(* IEC 61131-3 sources: Lasal-MCP/examples/SampleSource/LASALScreenAdvancedSolution/LASALScreenAdvancedSolution/LASALScreenAdvacnedSolution/Stations/Terminal/HMI/Network/DragDropNet, 1 file *)

(* ---- ONE_DragDropNet_Table.st ---- *)
#define OBJECTS_CONFIG

FUNCTION GLOBAL TAB ONE_DragDropNet
-1$UINT, 0$UINT,
0$UINT, 0$UINT,

6$UDINT,
TO_UDINT(2980745877), "_MyIO", 0$UINT, 3$UINT, 0$UINT,
TO_UDINT(3043040051), "_ScrollArea", 0$UINT, 15$UINT, 0$UINT,
TO_UDINT(2779823616), "_ScrollArea2", 0$UINT, 8$UINT, 0$UINT,
TO_UDINT(3157024878), "DragDropArea", 0$UINT, 0$UINT, 1$UINT,
TO_UDINT(1327562611), "IconDestList", 0$UINT, 0$UINT, 1$UINT,
TO_UDINT(1217922961), "IconSourceList", 0$UINT, 0$UINT, 1$UINT,

_NO_ATTR, TO_UDINT(694849416), "DRAGDROPAREA1",

_NO_ATTR, TO_UDINT(1251995598), "ICONDESTLIST1",

_NO_ATTR, TO_UDINT(77386850), "ICONSOURCELIST1",

//Internal connections
0$UDINT,
0$UDINT,
0$UDINT,
3$UDINT,
TO_UDINT(1), "DragDropArea", TO_UDINT(0), "Server0",
TO_UDINT(2), "DestList", TO_UDINT(1), "Server0",
TO_UDINT(2), "DragDropArea", TO_UDINT(0), "Server0",

//Initialization values
0$UDINT,
6$UDINT,
TO_UDINT(1), "VerticalLevel", TO_UDINT(1),//|DragDropNet.IconDestList1.VerticalLevel;
TO_UDINT(1), "LineWidth", TO_UDINT(100),//|DragDropNet.IconDestList1.LineWidth;
TO_UDINT(1), "ExtendedScrollBar", TO_UDINT(0),//|DragDropNet.IconDestList1.ExtendedScrollBar;
TO_UDINT(2), "VerticalLevel", TO_UDINT(1),//|DragDropNet.IconSourceList1.VerticalLevel;
TO_UDINT(2), "LineWidth", TO_UDINT(100),//|DragDropNet.IconSourceList1.LineWidth;
TO_UDINT(2), "ExtendedScrollBar", TO_UDINT(0),//|DragDropNet.IconSourceList1.ExtendedScrollBar;

//Symbolic initialization values
0$UDINT,
0$UDINT,

//Initialization of string values
0$UDINT,
0$UDINT,

//Configuration of tasks (RealTime, Cyclic, Background)
0$UDINT,
0$UDINT,

0$UDINT,
0$UDINT,

0$UDINT,
0$UDINT,

//External connections
0$UDINT,
3$UDINT,
TO_UDINT(0), "Lse", C_DIR, TO_UDINT(299963966), "Lse","Lse",
TO_UDINT(1), "Lse", C_DIR, TO_UDINT(299963966), "Lse","Lse",
TO_UDINT(2), "Lse", C_DIR, TO_UDINT(299963966), "Lse","Lse",

//Magic internal connections
0$UDINT,
0$UDINT,

//Configuration of timeslots of tasks (RealTime, Cyclic)
#ifdef __LSLLDR_TIMESLOTS__
0$UDINT,
0$UDINT,

0$UDINT,
0$UDINT,

#endif //__LSLLDR_TIMESLOTS__

//MultiMaster connections
#ifdef __LSLLDR_MULTIMASTER__
0$UDINT,
0$UDINT,
#endif //__LSLLDR_MULTIMASTER__

//Configuration for task ID (RealTime, CyclicTime)
#ifdef __LSLLDR_TASKID__
"\\\\TASKS2  "
0$UDINT,
0$UDINT,

0$UDINT,
0$UDINT,

0$UDINT,
0$UDINT,

#endif //__LSLLDR_TASKID__

END_FUNCTION
